// TIA Portal V19 export
TYPE "EM01_Output"
   STRUCT
      Status { S7_SetPoint := 'True'} : "EM_Output";
      BlowingActive : Bool;
      CalandriaActive : Bool;   // VÃ¡lvula proporcional de calandria con apertura > 0 %
   END_STRUCT;
END_TYPE
